(* IEC 61131-3 sources: codesys-framework/txt/application/WeVe Utils (library)/TimeStamp/DUT, 2 files *)

(* ---- E_TimeBase.dut.st ---- *)
{attribute 'qualified_only'}
{attribute 'strict'}
TYPE E_TimeBase :
(
	NTP 	:= 0,
	Manual 	:= 2
);
END_TYPE

(* ---- E_TimeZone.dut.st ---- *)
{attribute 'qualified_only'}
{attribute 'strict'}
TYPE E_TimeZone :
(
	Unknown							:=	0,
	GST_Dubai_UTC_4					:=	2,
	AFT_Kabul_UTC_4_30				:=	3,
	ART_Buenos_Aires_UTC_3			:=	19,
	AEDT_Melbourne_UTC_11			:=	37,
	AEST_Brisbane_UTC_10			:=	40,
	ACDT_Adelaide_UTC_10_30			:=	42,
	ACST_Darwin_UTC_9_30			:=	43,
	ACWST_Eucla_UTC_8_45			:=	45,
	BST_Dhaka_UTC_6					:=	51,
	CET_CEST_Brussels_UTC_1_2		:=	52,
	NST_St_Johns_UTC_3_30			:=	84,
	MST_Calgary_UTC_7				:=	102,
	CST_Beijing_UTC_8				:=	124,
	CVT_Praia_UTC_1					:=	129,
	EET_Cairo_UTC_2					:=	145,
	GMT_London_UTC_0				:=	161,
	GST_King_Edward_Point_UTC_2		:=	177,
	WIB_Jakarta_UTC_7				:=	187,
	IST_New_Delhi_UTC_5_30			:=	194,
	JST_Tokyo_UTC_9					:=	203,
	LINT_Kiritimati_UTC_14			:=	209,
	MMT_Rangoon_UTC_6_30			:=	243,
	NPT_Kathmandu_UTC_5_45			:=	278,
	NUT_Alofi_UTC_11				:=	280,
	NZDT_Auckland_UTC_13			:=	281,
	CHADT_Chatham_Islands_UTC_13_45	:=	282,
	MART_Taiohae_UTC_9_30			:=	287,
	MSK_Moscow_UTC_3				:=	309,
	ANAT_Anadyr_UTC_12				:=	334,
	EST_New_York_UTC_5				:=	379,
	PST_Los_Angeles_UTC_8			:=	399,
	HST_Honolulu_UTC_10				:=	407,
	UZT_Tashkent_UTC_5				:=	410,
	VET_Caracas_UTC_4				:=	413

);
END_TYPE
